//Raw diagnostic bytes; preserves existing high-byte-first order.
TYPE ST_DiagnosticElementRawIn :
STRUCT
    nHigh: ST_8Bit; //Diagnostic bits 8..15: pulse-test error and inputs 1..4.
    nLow: ST_8Bit; //Diagnostic bits 0..7: element status and errors.
END_STRUCT
END_TYPE

(* stored: Version 1.1.0.1
   DUT ST_DiagnosticElementRawIn: Id {73f839cd-bda8-090a-1863-d7a20736ae01} *)
